(* IEC 61131-3 sources: rusty/tests/lit/single/type_promotion/implicit_conversion, 2 files *)

(* ---- conversions_are_silent.st ---- *)
// RUN: %COMPILE %s 2> %t.err && %RUN | %CHECK %s
// RUN: not grep -E "Implicit conversion from|Operand of type" %t.err
// Explicit conversions, standard date and time arithmetic, builtins, generics and compiler-generated code
// never report an implicit conversion.
INTERFACE Source
    METHOD next : UDINT END_METHOD
END_INTERFACE

FUNCTION_BLOCK Counter IMPLEMENTS Source
    VAR count : UDINT; END_VAR
    METHOD next : UDINT
        count := count + 1;
        next := count;
    END_METHOD
END_FUNCTION_BLOCK

FUNCTION_BLOCK Wide EXTENDS Counter
END_FUNCTION_BLOCK

FUNCTION greeting : STRING
    greeting := 'hello';
END_FUNCTION

FUNCTION main
    VAR
        vSint : SINT := -3;
        vDint : DINT := 5;
        vLint : LINT := 6;
        vUdint : UDINT := 7;
        vUlint : ULINT := 8;
        vReal : REAL := 2.5;
        vTime : TIME := T#1s;
        vTod : TOD := TOD#01:00:00;
        vDt : DT := DT#2020-01-01-00:00:00;
        vDate : DATE := D#2020-01-02;
        counter : Counter;
        wide : Wide;
        source : Source;
        text : STRING;
    END_VAR

    // explicit conversions
    vUdint := TO_UDINT(vDint);
    vUlint := TO_ULINT(vLint);
    vReal := TO_REAL(vDint);
    vLint := TO_LINT(vReal);
    printf('%u %lu %f %ld$N', vUdint, vUlint, vReal, vLint);   // CHECK: 5 6 5.000000 5

    // counting idioms
    vUdint := vUdint + 1;
    vUdint := vUdint * 2;
    vUdint := vUdint - 1;
    printf('%u$N', vUdint);                                    // CHECK: 11

    // date and time arithmetic of the standard
    vTime := vTime + vTime;
    vTod := vTod + vTime;
    vDt := vDt + vTime;
    vTime := vDate - vDate;
    IF vTime = T#0s THEN
        printf('zero$N');                                      // CHECK: zero
    END_IF

    // generics and builtins
    vUdint := MAX(vUdint, vUdint);
    vUdint := SEL(TRUE, vUdint, 5);
    printf('%u$N', vUdint);                                    // CHECK: 5

    // generated code: constructors, vtables, aggregate returns, interface calls
    source := counter;
    vUdint := source.next();
    vUdint := wide.next();
    text := greeting();
    printf('%u %s$N', vUdint, text);                           // CHECK: 1 hello
END_FUNCTION

(* ---- sign_change_warnings.st ---- *)
// RUN: %PLC --check --error-format clang %s 2>&1 | %CHECK %s
// Implicit conversions that change the sign are reported where lowering has already rewritten the call.
FUNCTION_BLOCK Adder
    METHOD plus : UDINT
        VAR_INPUT amount : UDINT; END_VAR
        plus := amount;
    END_METHOD
END_FUNCTION_BLOCK

FUNCTION_BLOCK Stepper
    VAR_INPUT step : UDINT; END_VAR
END_FUNCTION_BLOCK

FUNCTION_BLOCK Producer
    VAR_OUTPUT out : DINT; END_VAR
END_FUNCTION_BLOCK

FUNCTION takesUdint : UDINT
    VAR_INPUT x : UDINT; END_VAR
    takesUdint := x;
END_FUNCTION

FUNCTION returnsUdint : UDINT
    VAR dint_ : DINT; END_VAR
    // CHECK: {{.*}}:[[@LINE+1]]:{{[0-9]+}}:{{.*}}warning[E160]: Implicit conversion from 'DINT' to 'UDINT' may change the sign.
    returnsUdint := dint_;
END_FUNCTION

FUNCTION main : DINT
    VAR
        adder : Adder;
        stepper : Stepper;
        producer : Producer;
        vDint : DINT;
        vUdint : UDINT;
        vUlint : ULINT;
        vLint : LINT;
        vByte : BYTE;
        vSint : SINT;
    END_VAR

    // CHECK: {{.*}}:[[@LINE+1]]:{{[0-9]+}}:{{.*}}warning[E160]: Implicit conversion from 'DINT' to 'UDINT' may change the sign.
    vUdint := vDint;
    // CHECK: {{.*}}:[[@LINE+1]]:{{[0-9]+}}:{{.*}}warning[E160]: Implicit conversion from 'LINT' to 'ULINT' may change the sign.
    vUlint := vLint;
    // CHECK: {{.*}}:[[@LINE+1]]:{{[0-9]+}}:{{.*}}warning[E160]: Implicit conversion from 'SINT' to 'BYTE' may change the sign.
    vByte := vSint;
    // CHECK: {{.*}}:[[@LINE+1]]:{{[0-9]+}}:{{.*}}warning[E160]: Implicit conversion from 'DINT' to 'UDINT' may change the sign.
    vUdint := takesUdint(vDint);
    // CHECK: {{.*}}:[[@LINE+1]]:{{[0-9]+}}:{{.*}}warning[E160]: Implicit conversion from 'DINT' to 'UDINT' may change the sign.
    vUdint := adder.plus(vDint);
    // CHECK: {{.*}}:[[@LINE+1]]:{{[0-9]+}}:{{.*}}warning[E160]: Implicit conversion from 'DINT' to 'UDINT' may change the sign.
    stepper(step := vDint);
    // CHECK: {{.*}}:[[@LINE+1]]:{{[0-9]+}}:{{.*}}warning[E160]: Implicit conversion from 'DINT' to 'UDINT' may change the sign.
    producer(out => vUdint);
    // CHECK: {{.*}}:[[@LINE+1]]:{{[0-9]+}}:{{.*}}warning[E161]: Operand of type 'UDINT' is converted to 'DINT', which may change its sign.
    vUdint := vUdint + vDint;
    // CHECK: {{.*}}:[[@LINE+1]]:{{[0-9]+}}:{{.*}}warning[E161]: Operand of type 'UDINT' is converted to 'DINT', which may change its sign.
    IF vDint < vUdint THEN
        vDint := 0;
    END_IF
END_FUNCTION
